FUNCTION_BLOCK logiBUS_ENC_ID (* Incremental encoder (quadrature A/B) as signed position *)
  (* Description: Copyright (c) 2026 HR Agrartechnik GmbH This program and the accompanying materials are made available under the terms of the Eclipse Public License 2.0 which is available at https://www.eclipse.org/legal/epl-2.0/ SPDX-License-Identifier: EPL-2.0 IN is the position as DINT in a DWORD (two's complement): convert it with DWORD_TO_DINT. Clockwise or counter-clockwise counts up depends on the wiring of A and B. Resolution: counts per quadrature cycle (4 edges). 1 = one count per detent for common rotary knobs, 4 = every edge. Other values are treated as 1. IND when the position changed, at most once per TimeRateLimit ms. TimeDelta > 0: additional IND every TimeDelta ms without change. RST sets the position to 0 and answers with CNF. The push button of a rotary knob is a normal digital input (Trainer20: Input_I9). *)
  (* Version 1.0, 2026-11-26, Franz Höpfinger, HR Agrartechnik GmbH, initial API and implementation and/or initial documentation *)
  PACKAGE logiBUS::io::ENC;
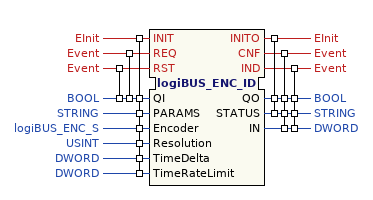
  EVENT_INPUT
    INIT : EInit WITH QI, PARAMS, Encoder, Resolution, TimeDelta, TimeRateLimit; (* Service Initialization *)
    REQ WITH QI; (* Service Request *)
    RST WITH QI; (* Set the position to 0 *)
  END_EVENT
  EVENT_OUTPUT
    INITO : EInit WITH QO, STATUS; (* Initialization Confirm *)
    CNF WITH QO, STATUS, IN; (* Confirmation of Requested Service *)
    IND WITH QO, STATUS, IN; (* Indication from Resource *)
  END_EVENT
  VAR_INPUT
    QI : BOOL; (* Event Input Qualifier *)
    PARAMS : STRING; (* Service Parameters *)
    Encoder : logiBUS::io::ENC::logiBUS_ENC_S := logiBUS_ENC::Invalid; (* Identify the encoder Encoder_E1 *)
    Resolution : USINT := 1; (* Counts per quadrature cycle: 1, 2 or 4 *)
    TimeDelta : DWORD; (* Additional IND every ms, 0 = only on change *)
    TimeRateLimit : DWORD := 50; (* Maximum 1 IND in how many ms (min. 10) *)
  END_VAR
  VAR_OUTPUT
    QO : BOOL; (* Event Output Qualifier *)
    STATUS : STRING; (* Service Status *)
    IN : DWORD; (* Position (DINT, convert with DWORD_TO_DINT) *)
  END_VAR
END_FUNCTION_BLOCK
